{attribute 'linkalways'} 
{attribute 'no_explicit_call' := 'This FB is a CLASS and must be accessed using methods or properties'}
{attribute 'enable_dynamic_creation'}
FUNCTION_BLOCK _ETcVnInterpolationType EXTENDS EnumDatatypeBase
VAR
	localData : ETcVnInterpolationType;
	activeData : REFERENCE TO ETcVnInterpolationType;
	enumBaseDatatype : _DINT(localData);
END_VAR

METHOD PRIVATE AddLocalEnumeration
VAR_INPUT
	Enumeration : T_MAXSTRING;
	Value : ETcVnInterpolationType;
END_VAR
AddEnumeration(Enumeration, Value);
END_METHOD

PROPERTY PUBLIC Address : PVOID
GET
Address := ADR(activeData);
END_GET
END_PROPERTY

METHOD PUBLIC ClearReference
VAR_INPUT
END_VAR
activeData REF= localData;
SetBaseDatatypeReference();
END_METHOD

METHOD PUBLIC Clone : I_Datatype
VAR
    pClone : POINTER TO _ETcVnInterpolationType;
END_VAR
pClone := __NEW(_ETcVnInterpolationType(InitialValue := Value));
Clone := pClone^;
END_METHOD

METHOD FB_init : BOOL
VAR_INPUT
	bInitRetains : BOOL; // if TRUE, the retain variables are initialized (warm start / cold start)
	bInCopyCode : BOOL;  // if TRUE, the instance afterwards gets moved into the copy code (online change)
	InitialValue : ETcVnInterpolationType;
END_VAR
localData := InitialValue;
AddBaseDatatype(enumBaseDatatype);
ClearReference();

AddLocalEnumeration('TCVN_IT_NEAREST_NEIGHBOR', ETcVnInterpolationType.TCVN_IT_NEAREST_NEIGHBOR);
AddLocalEnumeration('TCVN_IT_BILINEAR', ETcVnInterpolationType.TCVN_IT_BILINEAR);
AddLocalEnumeration('TCVN_IT_BICUBIC', ETcVnInterpolationType.TCVN_IT_BICUBIC);
AddLocalEnumeration('TCVN_IT_AREA_BASED', ETcVnInterpolationType.TCVN_IT_AREA_BASED);
AddLocalEnumeration('TCVN_IT_LANCZOS4', ETcVnInterpolationType.TCVN_IT_LANCZOS4);
AddLocalEnumeration('TCVN_IT_BILINEAR_EXACT', ETcVnInterpolationType.TCVN_IT_BILINEAR_EXACT);
AddLocalEnumeration('TCVN_IT_NEAREST_NEIGHBOR_EXACT', ETcVnInterpolationType.TCVN_IT_NEAREST_NEIGHBOR_EXACT);
END_METHOD

PROPERTY PUBLIC Identifier : T_MAXSTRING
GET
Identifier := 'ETcVnInterpolationType';
END_GET
END_PROPERTY

METHOD IsEnumeratorValueEqual : BOOL
VAR_INPUT
	Enumerator : I_KeyValueForwardEnumerator;
END_VAR
VAR
	storedValue : ETcVnInterpolationType;
END_VAR
IF NOT Enumerator.TryGet(storedValue) THEN
	RETURN;
END_IF

IsEnumeratorValueEqual := storedValue = activeData;
END_METHOD

METHOD PUBLIC MakeReferenceTo
VAR_INPUT
	ReferenceTarget : REFERENCE TO ETcVnInterpolationType;
END_VAR
activeData REF= ReferenceTarget;
SetBaseDatatypeReference();
END_METHOD

METHOD PROTECTED SetBaseDatatypeReference
VAR_INPUT
END_VAR
enumBaseDatatype.MakeReferenceTo(activeData);
END_METHOD

PROPERTY PUBLIC Size : UDINT
GET
Size := SIZEOF(activeData);
END_GET
END_PROPERTY

METHOD TryMakeReferenceTo : BOOL
VAR_INPUT
	Target : I_Datatype;
END_VAR
VAR
	pTargetData : POINTER TO ETcVnInterpolationType;
END_VAR
IF NOT IsEquivalentTo(Target) THEN
	RETURN;
END_IF

pTargetData := Target.Address;
activeData REF= pTargetData^;
SetBaseDatatypeReference();
TryMakeReferenceTo := TRUE;
END_METHOD

PROPERTY PUBLIC Value : ETcVnInterpolationType
GET
Value := activeData;
END_GET
SET
activeData := Value;
END_SET
END_PROPERTY

END_FUNCTION_BLOCK

(* stored: Version 1.1.0.1, ProductVersion 3.1.4024.13
   POU _ETcVnInterpolationType: Id {ba9e75ea-42dd-0bba-233c-e8fdd72b7315}, SpecialFunc None
   Folder Core: Id {2e742ac4-c5a2-00e6-18f2-a486752341d5}
   Folder Protected: Id {1febac23-bc12-0e7f-359d-2953f0ce94f8}
   Folder Customize: Id {fb13efc1-560d-0be6-1be0-ffdec6d26e34}
   Folder Constructor: Id {a2ff181c-f51e-0479-348a-e32c0d30ae23}
   Folder Private: Id {961f7734-5d31-09b1-3480-324fad025a32}
   Folder Protected: Id {bf471ec0-62d3-0704-05f2-765715c5bf74}
   Method AddLocalEnumeration: Id {c52ca102-bfe5-07b9-1f0f-1b385daa1fec}
   Property Address: Id {b346fbac-3367-0077-26e5-50b612e41e90}
   Get Get: Id {2c459276-eb79-04dd-35af-7597a9b0e8dc}
   Method ClearReference: Id {21908c4d-8b16-0412-3652-33423548e991}
   Method Clone: Id {3c68b57b-e257-0887-0db6-d00ba9f9a5c2}
   Method FB_init: Id {90e6fcdb-3b53-0644-35b4-51f2e1bb969c}
   Property Identifier: Id {c2ac3934-f58a-015c-19a8-f155e14a13da}
   Get Get: Id {39b3ba09-cd88-08a5-050f-0a240e2f6694}
   Method IsEnumeratorValueEqual: Id {19d17fe2-2b7d-0e09-3445-a3de39075fe9}
   Method MakeReferenceTo: Id {5a39876c-d73c-0800-074d-07a171eca940}
   Method SetBaseDatatypeReference: Id {8e36b850-ce3f-042c-30d0-9f291c5a906f}
   Property Size: Id {881580f5-cf13-0a05-2526-0dec540b5cc1}
   Get Get: Id {e7c48a3d-b75e-0181-00ba-393d13c55d86}
   Method TryMakeReferenceTo: Id {0070a147-d899-0157-3023-ed6c565d9c8a}
   Property Value: Id {662a6ce0-39e8-0e0d-2616-1e054740c6bd}
   Get Get: Id {121c3126-750d-02b1-02c6-0edc3f72b472}
   Set Set: Id {bf453bde-a1bb-025e-3b7d-10af8115e3d8} *)
